FUNCTION_BLOCK Sorting (* The equipment overview; the operator interface is internal to Control. *)
  (* Standard: 61499-2 *)
  (* Version 3.0, 2026-11-12, sorting2n, sorting2n, Complete hierarchical architecture with preserved leaf behavior *)
  PACKAGE Main;
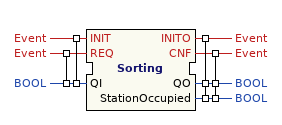
  EVENT_INPUT
    INIT WITH QI;
    REQ WITH QI;
  END_EVENT
  EVENT_OUTPUT
    INITO WITH QO, StationOccupied;
    CNF WITH QO, StationOccupied;
  END_EVENT
  VAR_INPUT
    QI : BOOL := FALSE;
  END_VAR
  VAR_OUTPUT
    QO : BOOL := FALSE;
    StationOccupied : BOOL := FALSE;
  END_VAR
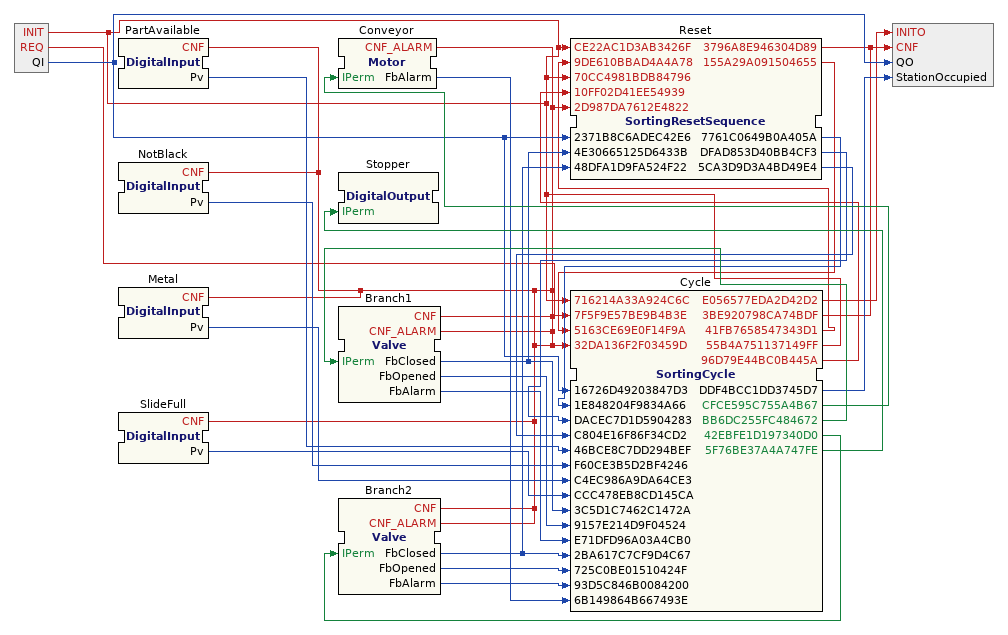
  FBS
    Conveyor : Motor; (* Move the part past the sensors *)
    Branch1 : Valve;
    Branch2 : Valve;
    Stopper : DigitalOutput;
    PartAvailable : DigitalInput;
    NotBlack : DigitalInput;
    Metal : DigitalInput;
    SlideFull : DigitalInput;
    Reset : SortingResetSequence; (* The complete three step conveyor reset. *)
    Cycle : SortingCycle; (* One minimal Reset / Run / Stop coordinator, movement procedures and equipment readiness. *)
  END_FBS
  EVENT_CONNECTIONS
    INIT TO Reset.CE22AC1D3AB3426F;
    INIT TO Cycle.716214A33A924C6C;
    REQ TO Cycle.7F5F9E57BE9B4B3E;
    Cycle.E056577EDA2D42D2 TO INITO;
    Cycle.3BE920798CA74BDF TO CNF;
    Reset.3796A8E946304D89 TO CNF;
    Cycle.41FB7658547343D1 TO Reset.9DE610BBAD4A4A78;
    Cycle.55B4A751137149FF TO Reset.70CC4981BDB84796;
    Cycle.55B4A751137149FF TO Reset.CE22AC1D3AB3426F;
    Cycle.96D79E44BC0B445A TO Reset.10FF02D41EE54939;
    Reset.155A29A091504655 TO Cycle.5163CE69E0F14F9A;
    PartAvailable.CNF TO Cycle.32DA136F2F03459D;
    NotBlack.CNF TO Cycle.32DA136F2F03459D;
    Metal.CNF TO Cycle.32DA136F2F03459D;
    SlideFull.CNF TO Cycle.32DA136F2F03459D;
    Branch1.CNF TO Cycle.32DA136F2F03459D;
    Branch1.CNF_ALARM TO Cycle.32DA136F2F03459D;
    Branch1.CNF TO Reset.2D987DA7612E4822;
    Branch2.CNF TO Cycle.32DA136F2F03459D;
    Branch2.CNF_ALARM TO Cycle.32DA136F2F03459D;
    Branch2.CNF TO Reset.2D987DA7612E4822;
    Conveyor.CNF_ALARM TO Cycle.32DA136F2F03459D;
  END_CONNECTIONS
  DATA_CONNECTIONS
    QI TO Reset.2371B8C6ADEC42E6;
    QI TO Cycle.16726D49203847D3;
    QI TO QO;
    Cycle.DDF4BCC1DD3745D7 TO StationOccupied;
    Reset.7761C0649B0A405A TO Cycle.1E848204F9834A66;
    Reset.DFAD853D40BB4CF3 TO Cycle.DACEC7D1D5904283;
    Reset.5CA3D9D3A4BD49E4 TO Cycle.C804E16F86F34CD2;
    PartAvailable.Pv TO Cycle.46BCE8C7DD294BEF;
    NotBlack.Pv TO Cycle.F60CE3B5D2BF4246;
    Metal.Pv TO Cycle.C4EC986A9DA64CE3;
    SlideFull.Pv TO Cycle.CCC478EB8CD145CA;
    Branch1.FbClosed TO Cycle.3C5D1C7462C1472A;
    Branch1.FbOpened TO Cycle.9157E214D9F04524;
    Branch1.FbAlarm TO Cycle.E71DFD96A03A4CB0;
    Branch1.FbClosed TO Reset.4E30665125D6433B;
    Branch2.FbClosed TO Cycle.2BA617C7CF9D4C67;
    Branch2.FbOpened TO Cycle.725C0BE01510424F;
    Branch2.FbAlarm TO Cycle.93D5C846B0084200;
    Branch2.FbClosed TO Reset.48DFA1D9FA524F22;
    Conveyor.FbAlarm TO Cycle.6B149864B667493E;
  END_CONNECTIONS
  ADAPTER_CONNECTIONS
    Cycle.CFCE595C755A4B67 TO Conveyor.IPerm;
    Cycle.BB6DC255FC484672 TO Branch1.IPerm;
    Cycle.42EBFE1D197340D0 TO Branch2.IPerm;
    Cycle.5F76BE37A4A747FE TO Stopper.IPerm;
  END_CONNECTIONS
END_FUNCTION_BLOCK
